Fanuc KAREL source: kt00700.KL

PROGRAM KT00700
%STACKSIZE=65535
%PRIORITY=65535
%NOLOCKGROUP
VAR
OUT : INTEGER
-- UNRESOLVED DECLARATIONS (source type spelling not recovered)
-- C1 : TYPE_0x001C (type_u16=0x001C)
-- C2 : TYPE_0x001C (type_u16=0x001C)
BEGIN
-- UNRESOLVED_PC line 8 opcodes [9D 22 A5] marker_code=0
-- UNRESOLVED_PC line 9 opcodes [9C 22 A5] marker_code=15
-- UNRESOLVED_PC line 10 opcodes [9D 22 A5] marker_code=30
-- UNRESOLVED_PC line 11 opcodes [9C 22 A5] marker_code=45
OUT=C1
END KT00700
